Staubli VAL3: Init.pgx

program Init()
  local num i
  local string l_sArmType
begin
  //dio

  //****************bool*****************
  _bEndCycle=false
  _bAtHome=false
  _bHeavyAlarm=false
  //判断是否是4轴机器人
  l_sArmType=left(getVersion("Arm Type"),2)
  _bIsScara=(l_sArmType=="rs" or l_sArmType=="ts" or l_sArmType=="tp")


  call rs:init()

end
